// Model of a two channel safe output terminal (EL2912): a TwinSAFE connection with two channels.
// Declare it in its group:  outputTerminal : T_SafeOutputTerminal2(group := safetyGroup);
// SafeOut1..2 are wired from FB outputs; Channel1..2 are the simulated field outputs,
// forced FALSE (fail-safe) unless the connection is in the Data state and the group is in RUN (OutputsEnabled).
FUNCTION_BLOCK T_SafeOutputTerminal2 EXTENDS T_SafeConnection
VAR_INPUT
    SafeOut1 : BOOL;
    SafeOut2 : BOOL;
END_VAR
VAR_OUTPUT
    Channel1 : BOOL;
    Channel2 : BOOL;
END_VAR

SUPER^();
Channel1 := SafeOut1 AND OutputsEnabled;
Channel2 := SafeOut2 AND OutputsEnabled;

END_FUNCTION_BLOCK

(* stored: Version 1.1.0.1
   POU T_SafeOutputTerminal2: Id {743b179f-a625-47bd-ad52-dc17aa13cae9}, SpecialFunc None *)
